Universal Robots PolyScope program: FeatureTest.urp

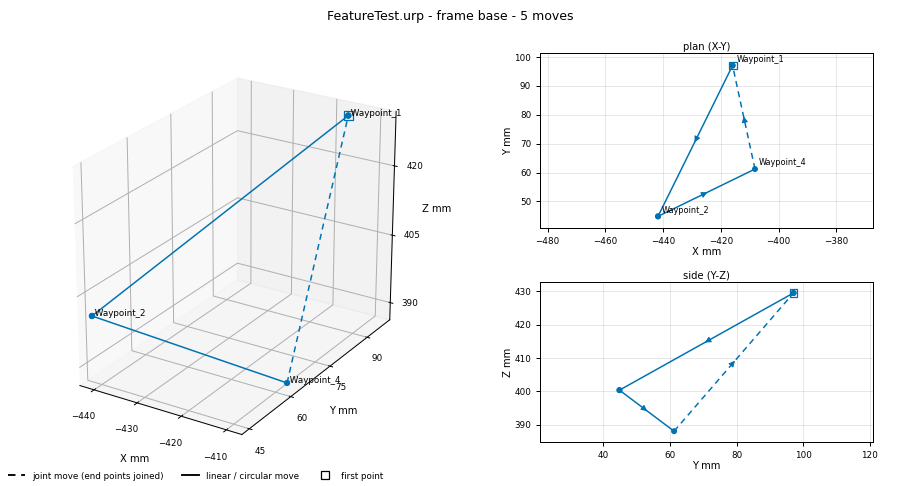
[picture p0: tool path of FeatureTest.urp in frame base, 5 of 5 moves have a stored position in this frame; points joined in program order, loops and branches not executed]
Program FeatureTest (createdIn=3.0.0 lastSavedIn=3.0.0 directory=/programs installation=default)
Robot Program (runOnlyOnce=true motionType=MoveJ speed=1.047198 acceleration=1.396263 useActiveTCP=false)
  'Program generated by VerticalBot Studio for UR5e on 25/10/2026 12:00:00'
  'Using nominal kinematics.'
  'Using Ref. Frame 2: p[0.100000, -0.050000, 0.020000, 0.000000, 0.000000, 0.523599]'
  'Using TCP Tool 1: p[0.010000, 0.000000, 0.120000, 0.000000, 0.261799, 0.000000]'
  Script: set_tcp(p[0.010000, 0.000000, 0.120000, 0.000000, 0.261799, 0.000000])
  Script: movej([-0.523599, -1.745329, 1.570796, -1.396263, -1.570796, 0.349066],6.98132,1.57080,0,0.0000)
  MoveJ speed 90.01 deg/s, acceleration 399.98 deg/s^2 (useActiveTCP=true)
    Waypoint Waypoint_1: TCP in base x=-415.957 y=97.082 z=429.557 mm, rx=-2.8465 ry=-1.036 rz=-0.3747 rad; joints [-30, -100, 90, -80, -90, 20] deg; flange x=-423.617 y=90.654 z=549.557 mm, rx=2.9521 ry=1.0745 rz=0 rad
  MoveL speed 300 mm/s, acceleration 1500 mm/s^2 (useActiveTCP=true)
    Waypoint Waypoint_2: motionParameters(blendRadius=0.005); TCP in base x=-441.769 y=44.852 z=400.392 mm, rx=-2.784 ry=-1.254 rz=-0.442 rad; joints [-22, -96, 90, -80, -90, 20] deg; flange x=-456.215 y=40.554 z=519.861 mm, rx=2.8233 ry=1.257 rz=0.075 rad
  'Circular move (R55.6 mm)'
  Script: movec(p[-0.408198, 0.061237, 0.388074, -2.843025, -1.166595, -0.465806],p[-0.414384, 0.147916, 0.407797, -2.938632, -0.908861, -0.436254],1.50000,0.30000,0.0050)
  MoveL speed 50 mm/s, acceleration 1500 mm/s^2 (useActiveTCP=true)
    Waypoint Waypoint_3: TCP in base x=-441.769 y=44.852 z=400.392 mm, rx=-2.784 ry=-1.254 rz=-0.442 rad; joints [-22, -96, 90, -80, -90, 20] deg; flange x=-456.215 y=40.554 z=519.861 mm, rx=2.8233 ry=1.257 rz=0.075 rad
  MoveL speed 300 mm/s, acceleration 1500 mm/s^2 (useActiveTCP=true)
    Waypoint Waypoint_4: TCP in base x=-408.198 y=61.237 z=388.074 mm, rx=-2.843 ry=-1.1666 rz=-0.4658 rad; joints [-26, -100, 95, -80, -90, 20] deg; flange x=-424.78 y=58.869 z=507.319 mm, rx=2.8515 ry=1.1521 rz=0.0898 rad
  Set DigitalOutput pin=digital_out[3]; digitalValue=1
  Set DigitalOutput pin=DO_GRIP; digitalValue=0
  Wait DigitalInput pin=digital_in[get_standard_digital_in(5)]; digitalValue=1
  Wait DigitalInput pin=DI_PART; digitalValue=1
  Wait Sleep waitTime=0.5
  'a comment line'
  Popup Message (haltProgram=false message=Hello operator)
  Call MyFunc
  Call SetRPM
  Script: RAW_CODE_LINE
  Call SubPick
  'Using TCP Tool 1: p[0.010000, 0.000000, 0.120000, 0.000000, 0.261799, 0.000000]'
  Script: set_tcp(p[0.010000, 0.000000, 0.120000, 0.000000, 0.261799, 0.000000])
  'Attach to Tool 1'
  Script: movej([-0.523599, -1.745329, 1.570796, -1.396263, -1.570796, 0.349066],6.98132,0.78540,0,0.0000)
  MoveJ speed 44.98 deg/s, acceleration 399.98 deg/s^2 (useActiveTCP=true)
    Waypoint Waypoint_5: TCP in base x=-415.957 y=97.082 z=429.557 mm, rx=-2.8465 ry=-1.036 rz=-0.3747 rad; joints [-30, -100, 90, -80, -90, 20] deg; flange x=-423.617 y=90.654 z=549.557 mm, rx=2.9521 ry=1.0745 rz=0 rad
  Halt
SubProgram  [hidden by the author, left out]
SubProgram  [hidden by the author, left out]
SubProgram  [hidden by the author, left out]
SubProgram MyFunc [hidden by the author, left out]
SubProgram SetRPM [hidden by the author, left out]
SubProgram SubPick [hidden by the author, left out]
